FUNCTION_BLOCK "FB_MotorControl"

VAR_INPUT
    Pressure_LOW : DINT;
END_VAR

VAR_OUTPUT
    Motor_Critical : BOOL;
END_VAR

VAR
    Threshold : DINT := 36464;
END_VAR

BEGIN

    IF NOT (Pressure_LOW < Threshold) THEN // MUTATED: COND_NEGATE
        Motor_Critical := TRUE;
    ELSE
        Motor_Critical := FALSE;
    END_IF;

END_FUNCTION_BLOCK
